(* IEC 61131-3 sources: plc-vscode/tests/st/all/trust-platform/crates/trust-runtime/tests/fixtures/oscat/core/src/14_memory_modules, 1 file *)

(* ---- tests.st ---- *)
TEST_PROGRAM oscat_logic_memory_helpers_behave
VAR
    Fifo16 : FIFO_16;
    Fifo32 : FIFO_32;
    Stack16 : STACK_16;
    Stack32 : STACK_32;
END_VAR

Fifo16(DIN := DWORD#0, E := TRUE, RD := FALSE, WD := FALSE, RST := TRUE);
ASSERT_TRUE(IN := Fifo16.EMPTY);
ASSERT_FALSE(IN := Fifo16.FULL);

Fifo16(DIN := DWORD#11, E := TRUE, RD := FALSE, WD := TRUE, RST := FALSE);
ASSERT_FALSE(IN := Fifo16.EMPTY);
ASSERT_FALSE(IN := Fifo16.FULL);

Fifo16(DIN := DWORD#22, E := TRUE, RD := FALSE, WD := TRUE, RST := FALSE);
Fifo16(DIN := DWORD#0, E := TRUE, RD := TRUE, WD := FALSE, RST := FALSE);
ASSERT_EQUAL(EXPECTED := DWORD#11, ACTUAL := Fifo16.DOUT);
ASSERT_FALSE(IN := Fifo16.EMPTY);

Fifo16(DIN := DWORD#0, E := TRUE, RD := TRUE, WD := FALSE, RST := FALSE);
ASSERT_EQUAL(EXPECTED := DWORD#22, ACTUAL := Fifo16.DOUT);
ASSERT_TRUE(IN := Fifo16.EMPTY);

Fifo32(DIN := DWORD#0, E := TRUE, RD := FALSE, WD := FALSE, RST := TRUE);
Fifo32(DIN := DWORD#33, E := TRUE, RD := FALSE, WD := TRUE, RST := FALSE);
Fifo32(DIN := DWORD#0, E := TRUE, RD := TRUE, WD := FALSE, RST := FALSE);
ASSERT_EQUAL(EXPECTED := DWORD#33, ACTUAL := Fifo32.DOUT);
ASSERT_TRUE(IN := Fifo32.EMPTY);

Stack16(DIN := DWORD#0, E := TRUE, RD := FALSE, WD := FALSE, RST := TRUE);
ASSERT_TRUE(IN := Stack16.EMPTY);

Stack16(DIN := DWORD#11, E := TRUE, RD := FALSE, WD := TRUE, RST := FALSE);
Stack16(DIN := DWORD#22, E := TRUE, RD := FALSE, WD := TRUE, RST := FALSE);
Stack16(DIN := DWORD#0, E := TRUE, RD := TRUE, WD := FALSE, RST := FALSE);
ASSERT_EQUAL(EXPECTED := DWORD#22, ACTUAL := Stack16.DOUT);
ASSERT_FALSE(IN := Stack16.EMPTY);

Stack16(DIN := DWORD#0, E := TRUE, RD := TRUE, WD := FALSE, RST := FALSE);
ASSERT_EQUAL(EXPECTED := DWORD#11, ACTUAL := Stack16.DOUT);
ASSERT_TRUE(IN := Stack16.EMPTY);

Stack32(DIN := DWORD#0, E := TRUE, RD := FALSE, WD := FALSE, RST := TRUE);
Stack32(DIN := DWORD#44, E := TRUE, RD := FALSE, WD := TRUE, RST := FALSE);
Stack32(DIN := DWORD#0, E := TRUE, RD := TRUE, WD := FALSE, RST := FALSE);
ASSERT_EQUAL(EXPECTED := DWORD#44, ACTUAL := Stack32.DOUT);
ASSERT_TRUE(IN := Stack32.EMPTY);
END_TEST_PROGRAM
